// TIA Portal V15.1 export
DATA_BLOCK "Par"   // DB1
{ S7_Optimized_Access := 'TRUE' }
VERSION : 0.1
// stored: AutoNumber false, MemoryReserve 100
   VAR RETAIN
      SP : Int := 700;   // HMI entry: Setpoint, 0.1 degC (C07b)
      HYST : Int := 50;   // HMI entry: Restart hysteresis, 0.1 degC (C07b)
      STG : Int := 100;   // HMI entry: 2nd stage below SP - STG, 0.1 degC (C07c)
      TStart : Time := T#2M;   // HMI entry: Max. time heat request -> RUN (C07f)
      TDrnOn : Time := T#3S;   // HMI entry: Scrubber high level before drain opens (C04)
      TDrnOff : Time := T#5S;   // HMI entry: Scrubber level gone before drain closes (C04)
      TDrnMax : Time := T#10M;   // HMI entry: Scrubber drain max. continuous open time (C04a)
      SP_V : Int := 700;   // Validated value used by the program (R-11)
      HYST_V : Int := 50;   // Validated value used by the program (R-11)
      STG_V : Int := 100;   // Validated value used by the program (R-11)
      TStart_V : Time := T#2M;   // Validated value used by the program (R-11)
      TDrnOn_V : Time := T#3S;   // Validated value used by the program (R-11)
      TDrnOff_V : Time := T#5S;   // Validated value used by the program (R-11)
      TDrnMax_V : Time := T#10M;   // Validated value used by the program (R-11)
   END_VAR
BEGIN
END_DATA_BLOCK
